FUNCTION_BLOCK MagazineCtrl (* Basic Function Block Type *)
  (* Standard: 61499-2 *)
  (* Version 0.0, 7/2/2026, Template *)
  PACKAGE Main;
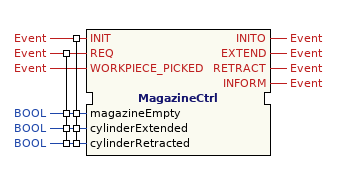
  EVENT_INPUT
    INIT WITH magazineEmpty, cylinderExtended, cylinderRetracted; (* Initialization Request *)
    REQ WITH magazineEmpty, cylinderExtended, cylinderRetracted; (* Normal Execution Request *)
    WORKPIECE_PICKED;
  END_EVENT
  EVENT_OUTPUT
    INITO; (* Initialization Confirm *)
    EXTEND; (* Execution Confirmation *)
    RETRACT;
    INFORM;
  END_EVENT
  VAR_INPUT
    magazineEmpty : BOOL; (* Input event qualifier *)
    cylinderExtended : BOOL;
    cylinderRetracted : BOOL;
  END_VAR
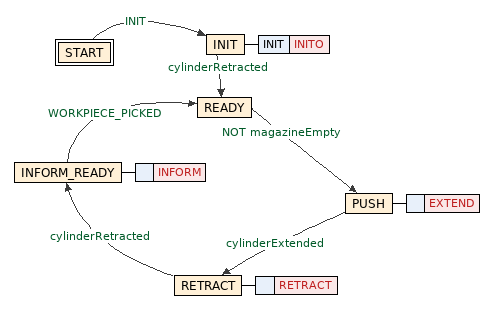
  EC_STATES
    START; (* Initial State *)
    INIT : INIT -> INITO; (* Initialization *)
    READY;
    PUSH : -> EXTEND;
    RETRACT : -> RETRACT;
    INFORM_READY : -> INFORM;
  END_STATES
  EC_TRANSITIONS
    START TO INIT := INIT;
    INIT TO READY := cylinderRetracted;
    READY TO PUSH := NOT magazineEmpty;
    PUSH TO RETRACT := cylinderExtended;
    RETRACT TO INFORM_READY := cylinderRetracted;
    INFORM_READY TO READY := WORKPIECE_PICKED;
  END_TRANSITIONS
  ALGORITHM INIT IN ST: (* Initialization algorithm *)
;
  END_ALGORITHM
  ALGORITHM REQ IN ST: (* Normally executed algorithm *)
;
  END_ALGORITHM
END_FUNCTION_BLOCK
